FUNCTION_BLOCK FB_Sensor
VAR_OUTPUT
	bActive	: BOOL;
END_VAR
VAR
	bSignal	AT %I*	: BOOL;
END_VAR

bActive := bSignal;

END_FUNCTION_BLOCK

(* stored: Version 1.1.0.1
   POU FB_Sensor: Id {8d408d6d-27ad-4505-bffa-752af12fe80f}, SpecialFunc None *)
